(* PLC project Motor_StartStop_TM241CE40T, PLCAutoPilot Machine Expert Logic Builder V19.2.3.0, author PLCAutoPilot *)
(* stored: creationDateTime 2025-12-30T21:00:00, version 1.0.0.0, modificationDateTime 2025-12-30T21:00:00 *)

PROGRAM PLC_PRG
  VAR
    EMERGENCY_PB AT %IX0.0 : BOOL;  (* Emergency Stop Push Button (NC - Normally Closed) *)
    START_PB AT %IX0.1 : BOOL;  (* Start Push Button (NO - Normally Open) *)
    STOP_PB AT %IX0.2 : BOOL;  (* Stop Push Button (NC - Normally Closed) *)
    MOTOR_OL AT %IX0.3 : BOOL;  (* Motor Overload Relay Contact (NC - Normally Closed) *)
    RESET_PB AT %IX0.4 : BOOL;  (* Alarm Reset Push Button (NO - Normally Open) *)
    MOTOR_RUN AT %QX0.0 : BOOL;  (* Motor Contactor Output *)
    MOTOR_LAMP AT %QX0.1 : BOOL;  (* Motor Running Indicator Lamp *)
    OL_ALARM_LAMP AT %QX0.2 : BOOL;  (* Overload Alarm Indicator Lamp *)
    READY_LAMP AT %QX0.3 : BOOL;  (* System Ready Indicator Lamp *)
    System_ready AT %M?0 : BOOL;  (* System Ready Flag - Set after 3 second startup delay *)
    Motor_sealed AT %M?1 : BOOL;  (* Motor Seal-in Memory Bit *)
    OL_Alarm_latched AT %M?2 : BOOL;  (* Overload Alarm Latched Memory Bit *)
  END_VAR
  VAR
    TON_Startup : TON;  (* 3 second startup delay timer *)
  END_VAR

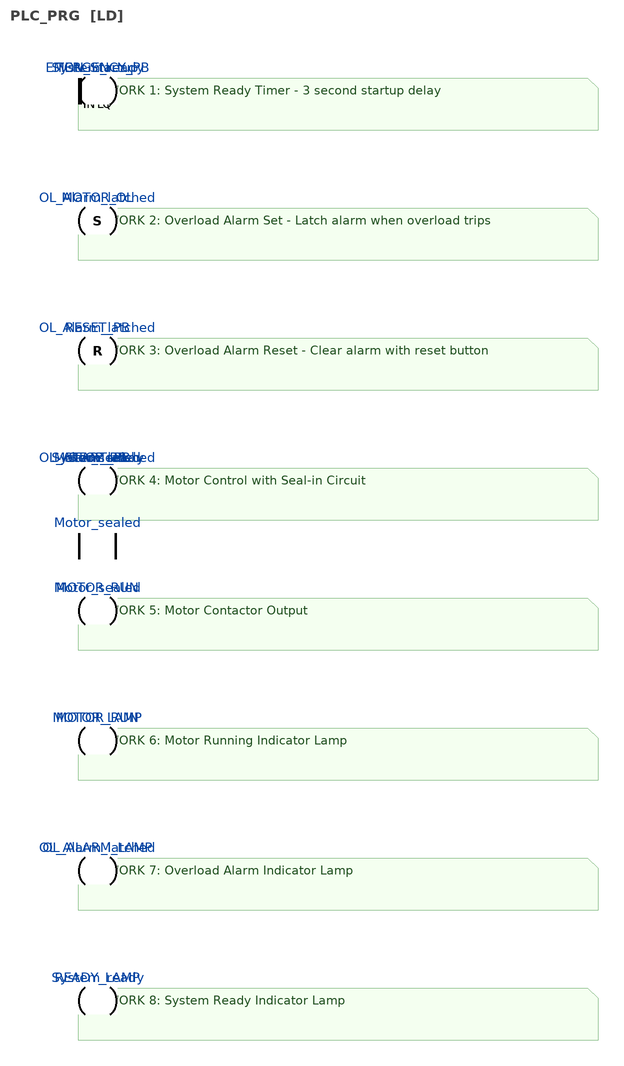
(* LD diagram, written out as Structured Text *)
(* NETWORK 1: System Ready Timer - 3 second startup delay *)
TON_Startup(IN := EMERGENCY_PB, PT := t#3s);
System_ready := TON_Startup.Q;
(* NETWORK 2: Overload Alarm Set - Latch alarm when overload trips *)
IF NOT MOTOR_OL THEN OL_Alarm_latched := TRUE; END_IF;
(* NETWORK 3: Overload Alarm Reset - Clear alarm with reset button *)
IF RESET_PB THEN OL_Alarm_latched := FALSE; END_IF;
(* NETWORK 4: Motor Control with Seal-in Circuit *)
Motor_sealed := System_ready AND (START_PB OR Motor_sealed) AND NOT STOP_PB AND NOT OL_Alarm_latched;
(* NETWORK 5: Motor Contactor Output *)
MOTOR_RUN := Motor_sealed;
(* NETWORK 6: Motor Running Indicator Lamp *)
MOTOR_LAMP := MOTOR_RUN;
(* NETWORK 7: Overload Alarm Indicator Lamp *)
OL_ALARM_LAMP := OL_Alarm_latched;
(* NETWORK 8: System Ready Indicator Lamp *)
READY_LAMP := System_ready;
END_PROGRAM
